FUNCTION_BLOCK StopAllMotion
VAR_INPUT
	
END_VAR
VAR_OUTPUT
END_VAR

VAR
	MotionState : INT;
	fbStopM1 : MC_Stop;
    fbStopM2 : MC_Stop;
    fbStopM3 : MC_Stop;
	fbHaltM1 : MC_Halt;
	fbHaltM2 : MC_Halt;
	fbHaltM3 : MC_Halt;
END_VAR

IF GVL_HMI.EmergencyStopIsOnHardware THEN
	MotionState := 10;  // Pressed Hardware Emergency Stop
	
ELSIF GVL_HMI.EmergencyStopIsOnSoftware THEN
	MotionState := 20;	// Pressed software Emergency Stop
	
ELSE
	MotionState := 30;	// Deactivation All STOPS
	
END_IF



CASE MotionState OF

10:	

    fbStopM1(
        Axis      := GVL_Axes.Axis1,
        Execute   := TRUE);   

    fbStopM2(
        Axis      := GVL_Axes.Axis2,
        Execute   := TRUE);

    fbStopM3(
        Axis      := GVL_Axes.Axis3,
        Execute   := TRUE);
	
20:	
    fbHaltM1(
        Axis      := GVL_Axes.Axis1,
        Execute   := TRUE);   

    fbHaltM2(
        Axis      := GVL_Axes.Axis2,
        Execute   := TRUE);

    fbHaltM3(
        Axis      := GVL_Axes.Axis3,
        Execute   := TRUE);
30: 

 fbStopM1(
        Axis      := GVL_Axes.Axis1,
        Execute   := FALSE);   

    fbStopM2(
        Axis      := GVL_Axes.Axis2,
        Execute   := FALSE);

    fbStopM3(
        Axis      := GVL_Axes.Axis3,
        Execute   := FALSE);


 fbHaltM1(
        Axis      := GVL_Axes.Axis1,
        Execute   := FALSE);   

    fbHaltM2(
        Axis      := GVL_Axes.Axis2,
        Execute   := FALSE);

    fbHaltM3(
        Axis      := GVL_Axes.Axis3,
        Execute   := FALSE);

	
END_CASE

END_FUNCTION_BLOCK

(* stored: Version 1.1.0.1, ProductVersion 3.1.4024.15
   POU StopAllMotion: Id {5fe55818-2cac-4d93-82ef-bf995b96a710}, SpecialFunc None *)
